TYPE E_SwitchEventType :
(
    ShortClick,
    LongClick,
    HoldStarted,
    HoldReleased
);
END_TYPE

(* stored: Version 1.1.0.1, ProductVersion 3.1.4026.20
   DUT E_SwitchEventType: Id {D1A10001-0A11-4A11-8A11-000000000001} *)
